Yaskawa INFORM job: SUBPICK.JBI

/JOB
//NAME SUBPICK
//POS
///NPOS 1,0,0,0,0,0
///TOOL 1
///POSTYPE PULSE
///PULSE
C00000=18,24,-10,30,-45,60
//INST
///DATE 2026/10/26 01:18
///COMM Generated using RoboDK
///ATTR SC,RW
///GROUP1 RB1
NOP
MOVL C00000 V=300.0 ACC=100 DEC=100
DOUT OT#(7) ON
END
